(* IEC 61131-3 sources: model-first-plc-agent-ai/results/T2-W-15, 2 files *)

(* ---- a1_code.st ---- *)
FUNCTION_BLOCK FillingRuntime
VAR_INPUT
    start : BOOL;
    stop : BOOL;
    LSH : BOOL;
    LSHH : BOOL;
    TimerDuration : TIME;
END_VAR
VAR_OUTPUT
    fill_valve : BOOL;
    discharge_valve : BOOL;
END_VAR
VAR
    ActiveState : INT := 0;
    PreviousState : INT;
    x0 : BOOL := TRUE;
    x1 : BOOL := FALSE;
    FillingTimer : TON;
    timer_done : BOOL := FALSE;
END_VAR

(* Evaluate the timer owned by the currently active filling step. *)
FillingTimer(IN := x1, PT := TimerDuration);
timer_done := FillingTimer.Q;

PreviousState := ActiveState;

CASE ActiveState OF
    0:
        IF start AND NOT stop AND NOT LSHH THEN
            ActiveState := 1;
        END_IF;

    1:
        IF stop OR LSHH OR timer_done THEN
            ActiveState := 0;
        END_IF;

ELSE
    ActiveState := 0;
END_CASE;

x0 := ActiveState = 0;
x1 := ActiveState = 1;

(* Start timing on entry and reset timing on exit. *)
IF ActiveState <> PreviousState THEN
    FillingTimer(IN := x1, PT := TimerDuration);
    timer_done := FALSE;
END_IF;

fill_valve := x1;
discharge_valve := FALSE;

END_FUNCTION_BLOCK

PROGRAM Main
VAR
    StartCommand AT %IX100.0 : BOOL;
    StopCommand AT %IX100.1 : BOOL;
    LSH AT %IX100.2 : BOOL;
    LSHH AT %IX100.3 : BOOL;
    FillValve AT %QX100.0 : BOOL;
    DischargeValve AT %QX100.1 : BOOL;
END_VAR
VAR
    (* Configure the required filling duration before operation. *)
    TimerDuration : TIME := T#0s;
    StartEdge : R_TRIG;
    RuntimeLogic : FillingRuntime;
END_VAR

StartEdge(CLK := StartCommand);

RuntimeLogic(
    start := StartEdge.Q,
    stop := StopCommand,
    LSH := LSH,
    LSHH := LSHH,
    TimerDuration := TimerDuration
);

FillValve := RuntimeLogic.fill_valve;
DischargeValve := RuntimeLogic.discharge_valve;

END_PROGRAM

(* ---- a2_code.st ---- *)
FUNCTION_BLOCK TankFillingController
VAR_INPUT
    StartCommand : BOOL;
    StopCommand : BOOL;
    LSH : BOOL;
    LSHH : BOOL;
    TimerDuration : TIME;
END_VAR
VAR_OUTPUT
    fill_valve : BOOL;
    discharge_valve : BOOL;
END_VAR
VAR
    StartEdge : R_TRIG;
    FillingTimer : TON;
    start : BOOL;
    stop : BOOL;
    timer_done : BOOL;
    x1 : BOOL := FALSE;
END_VAR

StartEdge(CLK := StartCommand);
start := StartEdge.Q;
stop := StopCommand;

IF stop THEN
    x1 := FALSE;
ELSIF NOT x1 AND start THEN
    x1 := TRUE;
END_IF;

FillingTimer(IN := x1, PT := TimerDuration);
timer_done := FillingTimer.Q;

IF x1 AND (stop OR LSHH OR timer_done) THEN
    x1 := FALSE;
    FillingTimer(IN := FALSE, PT := TimerDuration);
    timer_done := FillingTimer.Q;
END_IF;

fill_valve := x1;
discharge_valve := FALSE;

END_FUNCTION_BLOCK

PROGRAM Main
VAR
    StartCommand AT %IX100.0 : BOOL;
    StopCommand AT %IX100.1 : BOOL;
    LSH AT %IX100.2 : BOOL;
    LSHH AT %IX100.3 : BOOL;
    FillValve AT %QX100.0 : BOOL;
    DischargeValve AT %QX100.1 : BOOL;
END_VAR
VAR
    TimerDuration : TIME := T#10s;
    Controller : TankFillingController;
END_VAR

Controller(
    StartCommand := StartCommand,
    StopCommand := StopCommand,
    LSH := LSH,
    LSHH := LSHH,
    TimerDuration := TimerDuration
);

FillValve := Controller.fill_valve;
DischargeValve := Controller.discharge_valve;

END_PROGRAM
